(* IEC 61131-3 sources: kns-port-domestic/tools/inventory_tests/fixtures/lib/src/GVLs, 1 file *)

(* ---- GVL_Lib.gvl.st ---- *)
{attribute 'qualified_only'}
// Константы и переменные в одном списке (для PLCopenXML так нельзя)
VAR_GLOBAL CONSTANT
    MAX_ITEMS : INT := 8;
END_VAR
VAR_GLOBAL
    {attribute 'symbol' := 'read'}
    iItems : INT;
END_VAR
